DATA_BLOCK "HMI ALARMS"
TITLE =HMI Alarms - NS12
//One BOOL per alarm, written by FC1220 every scan (no latching here: the
//fault bits keep their own latch / reset). NS12 address: SERIALA:DB0013_DBXbbbbb.ii
//v1.1 2026-11-24: DBX9.6 Any_Fault (bytes 0...8) and DBX9.7 Any_Alarm (+ status
//9.0...9.3) for the NS12 alarm bar Control Flag (bar shown only when needed).
VERSION : 1.1


  STRUCT
   Fuse_Fault : BOOL ;	//DBX0.0 Fuse fault
   Motor_Protect : BOOL ;	//DBX0.1 Motor protection tripped
   Motor_Temp : BOOL ;	//DBX0.2 Motor temperature fault
   Air_Low : BOOL ;	//DBX0.3 Compressed air below 5 bar
   EStop_Desk_X120 : BOOL ;	//DBX0.4 E-STOP desk X120 (HMI box)
   EStop_Desk_X121 : BOOL ;	//DBX0.5 E-STOP desk X121 (feeder box)
   EStop_Elevator : BOOL ;	//DBX0.6 E-STOP elevator station
   EStop_Flipper : BOOL ;	//DBX0.7 E-STOP flipper station
   Door_Feeder : BOOL ;	//DBX1.0 Door open - feeder
   Door_Elevator : BOOL ;	//DBX1.1 Door open - elevator
   Door_Flipper : BOOL ;	//DBX1.2 Door open - flipper
   Spare_1_3 : BOOL ;	//DBX1.3 Spare
   Spare_1_4 : BOOL ;	//DBX1.4 Spare
   Spare_1_5 : BOOL ;	//DBX1.5 Spare
   Spare_1_6 : BOOL ;	//DBX1.6 Spare
   Spare_1_7 : BOOL ;	//DBX1.7 Spare
   C2_Angle_Fault : BOOL ;	//DBX2.0 C2 angle conveyor fault
   Elev_Rollers_Fault : BOOL ;	//DBX2.1 Elevator rollers (C0) fault
   Elev_Pusher_Fault : BOOL ;	//DBX2.2 Elevator pusher fault
   Elev_Not_Centered : BOOL ;	//DBX2.3 Elevator - packet not centered
   C4_Fault : BOOL ;	//DBX2.4 C4 collator fault
   C4_Timeout : BOOL ;	//DBX2.5 C4 collator timeout stop
   C4_Infeed_Obstruct : BOOL ;	//DBX2.6 C4 infeed obstruction
   C6_Fault : BOOL ;	//DBX2.7 C6 flipper delivery fault
   Flipper_Obstruct : BOOL ;	//DBX3.0 Flipper flip obstructed
   C10_Fault : BOOL ;	//DBX3.1 C10 pivot conveyor fault
   Pivot_Timeout : BOOL ;	//DBX3.2 Pivot timeout
   Pivot_Conflict : BOOL ;	//DBX3.3 Pivot / conveyor conflict
   C13_Delivery_Fault : BOOL ;	//DBX3.4 C13 delivery fault (low)
   C23_Delivery_Fault : BOOL ;	//DBX3.5 C23 delivery fault (high)
   Spare_3_6 : BOOL ;	//DBX3.6 Spare
   Spare_3_7 : BOOL ;	//DBX3.7 Spare
   VFD_U44_3 : BOOL ;	//DBX4.0 Drive U44.3 fault - C4
   VFD_U45_0 : BOOL ;	//DBX4.1 Drive U45.0 fault - C5
   VFD_U45_3 : BOOL ;	//DBX4.2 Drive U45.3 fault - C6
   VFD_U45_6 : BOOL ;	//DBX4.3 Drive U45.6 fault - C7 flipper conveyor
   VFD_U46_0 : BOOL ;	//DBX4.4 Drive U46.0 fault - Flipper
   VFD_U46_4 : BOOL ;	//DBX4.5 Drive U46.4 fault - C8 turntable conveyor
   VFD_U47_0 : BOOL ;	//DBX4.6 Drive U47.0 fault - Turntable
   VFD_U47_5 : BOOL ;	//DBX4.7 Drive U47.5 fault - C9 pusher 2 conveyor
   VFD_U47_6 : BOOL ;	//DBX5.0 Drive U47.6 fault - Pusher 2
   VFD_U48_0 : BOOL ;	//DBX5.1 Drive U48.0 fault - C10
   VFD_U48_3 : BOOL ;	//DBX5.2 Drive U48.3 fault - C11
   VFD_U48_6 : BOOL ;	//DBX5.3 Drive U48.6 fault - C12
   VFD_U49_0 : BOOL ;	//DBX5.4 Drive U49.0 fault - C13
   VFD_U53_2 : BOOL ;	//DBX5.5 Drive U53.2 fault - C21
   VFD_U53_4 : BOOL ;	//DBX5.6 Drive U53.4 fault - C22
   VFD_U54_0 : BOOL ;	//DBX5.7 Drive U54.0 fault - C23
   Sens_B5_1_On : BOOL ;	//DBX6.0 Sensor Elevator platform infeed B5.1 ON - line empty (packet left or dir
   Sens_B5_2_On : BOOL ;	//DBX6.1 Sensor Elevator platform limit B5.2 ON - line empty (packet left or dirt
   Sens_B5_4_On : BOOL ;	//DBX6.2 Sensor C1 exit B5.4 ON - line empty (packet left or dirty sensor)
   Sens_B5_5_On : BOOL ;	//DBX6.3 Sensor C2 infeed B5.5 ON - line empty (packet left or dirty sensor)
   Sens_B6_0_On : BOOL ;	//DBX6.4 Sensor C2 roller center B6.0 ON - line empty (packet left or dirty senso
   Sens_B6_7_On : BOOL ;	//DBX6.5 Sensor C4 infeed B6.7 ON - line empty (packet left or dirty sensor)
   Sens_B7_0_On : BOOL ;	//DBX6.6 Sensor C4 exit B7.0 ON - line empty (packet left or dirty sensor)
   Sens_B7_1_On : BOOL ;	//DBX6.7 Sensor C5 exit B7.1 ON - line empty (packet left or dirty sensor)
   Sens_B7_2_On : BOOL ;	//DBX7.0 Sensor C6 reaching B7.2 ON - line empty (packet left or dirty sensor)
   Sens_B7_3_On : BOOL ;	//DBX7.1 Sensor C6 exit B7.3 ON - line empty (packet left or dirty sensor)
   Sens_B7_4_On : BOOL ;	//DBX7.2 Sensor Flipper infeed B7.4 ON - line empty (packet left or dirty sensor)
   Sens_B8_2_On : BOOL ;	//DBX7.3 Sensor Flipper exit B8.2 ON - line empty (packet left or dirty sensor)
   Sens_B9_6_On : BOOL ;	//DBX7.4 Sensor C9 infeed B9.6 ON - line empty (packet left or dirty sensor)
   Sens_B9_7_On : BOOL ;	//DBX7.5 Sensor C9 packet edge B9.7 ON - line empty (packet left or dirty sensor)
   Sens_B10_4_On : BOOL ;	//DBX7.6 Sensor C10 infeed B10.4 ON - line empty (packet left or dirty sensor)
   Sens_B10_5_On : BOOL ;	//DBX7.7 Sensor C10 full B10.5 ON - line empty (packet left or dirty sensor)
   Sens_B10_7_On : BOOL ;	//DBX8.0 Sensor C11 exit B10.7 ON - line empty (packet left or dirty sensor)
   Sens_B11_0_On : BOOL ;	//DBX8.1 Sensor C12 exit B11.0 ON - line empty (packet left or dirty sensor)
   Sens_B11_1_On : BOOL ;	//DBX8.2 Sensor C13 slow B11.1 ON - line empty (packet left or dirty sensor)
   Sens_B5_4_Off : BOOL ;	//DBX8.3 Sensor C1 exit B5.4 OFF - line empty (check sensor / reflector)
   Sens_B9_7_Off : BOOL ;	//DBX8.4 Sensor C9 packet edge B9.7 OFF - line empty (check sensor / reflector)
   Spare_8_5 : BOOL ;	//DBX8.5 Spare
   Spare_8_6 : BOOL ;	//DBX8.6 Spare
   Spare_8_7 : BOOL ;	//DBX8.7 Spare
   Clearing_Active : BOOL ;	//DBX9.0 Clearing (F4) active
   Packets_Present : BOOL ;	//DBX9.1 Packets present on C1-C2 / C7-C9
   Control_Off : BOOL ;	//DBX9.2 Control voltage OFF - press START
   Start_Ready : BOOL ;	//DBX9.3 Start ready (10 s)
   Spare_9_4 : BOOL ;	//DBX9.4 Spare
   Spare_9_5 : BOOL ;	//DBX9.5 Spare
   Any_Fault : BOOL ;	//DBX9.6 At Least One Fault (DBX0.0...8.7) - NS12 Alarm Bar Display
   Any_Alarm : BOOL ;	//DBX9.7 At Least One Fault or Status Message (DBX0.0...9.3)
  END_STRUCT ;
BEGIN
   Fuse_Fault := FALSE;
   Motor_Protect := FALSE;
   Motor_Temp := FALSE;
   Air_Low := FALSE;
   EStop_Desk_X120 := FALSE;
   EStop_Desk_X121 := FALSE;
   EStop_Elevator := FALSE;
   EStop_Flipper := FALSE;
   Door_Feeder := FALSE;
   Door_Elevator := FALSE;
   Door_Flipper := FALSE;
   Spare_1_3 := FALSE;
   Spare_1_4 := FALSE;
   Spare_1_5 := FALSE;
   Spare_1_6 := FALSE;
   Spare_1_7 := FALSE;
   C2_Angle_Fault := FALSE;
   Elev_Rollers_Fault := FALSE;
   Elev_Pusher_Fault := FALSE;
   Elev_Not_Centered := FALSE;
   C4_Fault := FALSE;
   C4_Timeout := FALSE;
   C4_Infeed_Obstruct := FALSE;
   C6_Fault := FALSE;
   Flipper_Obstruct := FALSE;
   C10_Fault := FALSE;
   Pivot_Timeout := FALSE;
   Pivot_Conflict := FALSE;
   C13_Delivery_Fault := FALSE;
   C23_Delivery_Fault := FALSE;
   Spare_3_6 := FALSE;
   Spare_3_7 := FALSE;
   VFD_U44_3 := FALSE;
   VFD_U45_0 := FALSE;
   VFD_U45_3 := FALSE;
   VFD_U45_6 := FALSE;
   VFD_U46_0 := FALSE;
   VFD_U46_4 := FALSE;
   VFD_U47_0 := FALSE;
   VFD_U47_5 := FALSE;
   VFD_U47_6 := FALSE;
   VFD_U48_0 := FALSE;
   VFD_U48_3 := FALSE;
   VFD_U48_6 := FALSE;
   VFD_U49_0 := FALSE;
   VFD_U53_2 := FALSE;
   VFD_U53_4 := FALSE;
   VFD_U54_0 := FALSE;
   Sens_B5_1_On := FALSE;
   Sens_B5_2_On := FALSE;
   Sens_B5_4_On := FALSE;
   Sens_B5_5_On := FALSE;
   Sens_B6_0_On := FALSE;
   Sens_B6_7_On := FALSE;
   Sens_B7_0_On := FALSE;
   Sens_B7_1_On := FALSE;
   Sens_B7_2_On := FALSE;
   Sens_B7_3_On := FALSE;
   Sens_B7_4_On := FALSE;
   Sens_B8_2_On := FALSE;
   Sens_B9_6_On := FALSE;
   Sens_B9_7_On := FALSE;
   Sens_B10_4_On := FALSE;
   Sens_B10_5_On := FALSE;
   Sens_B10_7_On := FALSE;
   Sens_B11_0_On := FALSE;
   Sens_B11_1_On := FALSE;
   Sens_B5_4_Off := FALSE;
   Sens_B9_7_Off := FALSE;
   Spare_8_5 := FALSE;
   Spare_8_6 := FALSE;
   Spare_8_7 := FALSE;
   Clearing_Active := FALSE;
   Packets_Present := FALSE;
   Control_Off := FALSE;
   Start_Ready := FALSE;
   Spare_9_4 := FALSE;
   Spare_9_5 := FALSE;
   Any_Fault := FALSE;
   Any_Alarm := FALSE;
END_DATA_BLOCK
